{attribute 'qualified_only'}
{attribute 'strict'}
{attribute 'to_string'}
TYPE E_PPStatus :
(
    UNKNOWN:= 0,
    IN := 1,
    OUT := 2
) UINT;
END_TYPE

(* stored: Version 1.1.0.1
   DUT E_PPStatus: Id {fdcd12af-97a1-4892-9e58-ae9e4d6b3612} *)
